FUNCTION_BLOCK AD2_TO_AD (* Composite FB for convert bidirectional AD2 to unidirectional AD *)
  (* Standard: 61499-2; Function: AD2_BIDIR forwards its incoming (EO1) side out as a plain unidirectional signal via AD_OUT. AD_IN publishes its value onto the outgoing (EI1) side of AD2_BIDIR.; Description: Copyright (c) 2026 HR Agrartechnik GmbH This program and the accompanying materials are made available under the terms of the Eclipse Public License 2.0 which is available at https://www.eclipse.org/legal/epl-2.0/ SPDX-License-Identifier: EPL-2.0 *)
  (* Version 1.0, 2026-11-13, Franz Höpfinger, HR Agrartechnik GmbH, Initial Version - Luecke geschlossen (analog zu AB2_TO_AB) *)
  PACKAGE adapter::conversion::bidirectional;
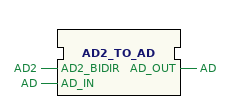
  SOCKETS
    AD2_BIDIR : adapter::types::bidirectional::AD2; (* Adapter Input: bidirectional tap, incoming side forwarded to AD_OUT, outgoing side driven by AD_IN *)
    AD_IN : adapter::types::unidirectional::AD; (* Adapter Input: unidirectional source *)
  END_SOCKETS
  PLUGS
    AD_OUT : adapter::types::unidirectional::AD; (* Adapter Output: mirrors AD2_BIDIR's incoming (indication) side *)
  END_PLUGS
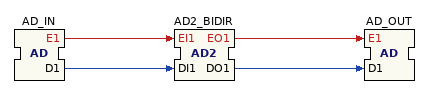
  EVENT_CONNECTIONS
    AD2_BIDIR.EO1 TO AD_OUT.E1;
    AD_IN.E1 TO AD2_BIDIR.EI1;
  END_CONNECTIONS
  DATA_CONNECTIONS
    AD2_BIDIR.DO1 TO AD_OUT.D1;
    AD_IN.D1 TO AD2_BIDIR.DI1;
  END_CONNECTIONS
END_FUNCTION_BLOCK
